PROGRAM MAIN
VAR
	{attribute 'OPC.UA.DA' := '1'}
	machine		: FB_Machine; //top-level module, start/stop with machine.ocmd
	
	(* Test harness
	----------------------------------------------------------------------------------------------------*)
	{attribute 'OPC.UA.DA' := '1'}
	softwareSim	: FB_ExampleSoftwareSim; //plays the software side of the station's trigger/tell
	{attribute 'OPC.UA.DA' := '1'}
	dosingSim	: FB_DosingProcessSim; //simulates the dosing station's flows
END_VAR

machine();

//Outside world: answers the example station's job requests
softwareSim(transaction := machine.exampleStation.transaction);

//Process simulation for the dosing station (turn off with dosingSim.cfg.enable when I/O is linked)
dosingSim(station := machine.dosingStation);

END_PROGRAM

(* stored: Version 1.1.0.1, ProductVersion 3.1.4024.12
   POU MAIN: Id {4db6d972-4f74-41c6-99a2-361264a8ef89}, SpecialFunc None *)
